SUBAPPLICATION Input_CLIENT_Method_IE (* logiBUS-Taster (logiBUS_IE) loest per CLIENT_0 einen argumentlosen OPC-UA-Methodenaufruf (CALL_METHOD) aus *)
  (* Standard: 61499-2; Description: Copyright (c) 2026 Meisterschulen am Ostbahnhof This program and the accompanying materials are made available under the terms of the Eclipse Public License 2.0 which is available at https://www.eclipse.org/legal/epl-2.0/ SPDX-License-Identifier: EPL-2.0 *)
  (* Version 1.1, 2026-10-18, Franz Höpfinger, Meisterschulen am Ostbahnhof, Wie Button_CLIENT_Method_IE, aber logiBUS_IE statt Button_IE (Taster statt VT-Button) *)
  (* Version 1.0, 2026-09-22, Franz Höpfinger, Meisterschulen am Ostbahnhof, initial implementation - herausgeloest aus logiBUS_AI_Calibrated_Subscribe_VT_OPC (Button_IE + CLIENT_0 kam dort 2x identisch vor, fuer CO und CS). Franz: 'Button_IE CLIENT_0 kann eine Subapp werden, das ist ein generelles Muster zum Rufen einer Methode vom VT aus' - InputEvent ist Parameter (nicht hartcodiert auf BT_PRESSED_LATCHED), damit auch andere Aktivierungsarten (z.B. Loslassen) wiederverwendbar sind. *)
  PACKAGE MyLib::sys;
  IMPORT logiBUS::io::DI::logiBUS_DI;
  IMPORT logiBUS::io::DI::logiBUS_DI_S;
  IMPORT logiBUS::io::DI::logiBUS_DI_Events_S;
  IMPORT logiBUS::io::DI::logiBUS_DI_Events::BUTTON_PRESS_DOWN;
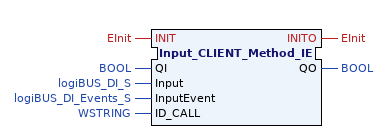
  EVENT_INPUT
    INIT : EInit; (* Initialization Request *)
  END_EVENT
  EVENT_OUTPUT
    INITO : EInit; (* Initialization Confirm *)
  END_EVENT
  VAR_INPUT
    QI : BOOL := TRUE; (* Quality Input - TRUE to enable service *)
    Input : logiBUS::io::DI::logiBUS_DI_S := logiBUS_DI::Invalid; (* Taster Input_I1..I8 *)
    InputEvent : logiBUS::io::DI::logiBUS_DI_Events_S := BUTTON_PRESS_DOWN; (* Welches Tasterereignis den Aufruf ausloest *)
    ID_CALL : WSTRING; (* Methodenadresse (ACTION=CALL_METHOD, mit Endpunkt, auch localhost) *)
  END_VAR
  VAR_OUTPUT
    QO : BOOL; (* Quality Output - TRUE if service executed successfully *)
  END_VAR
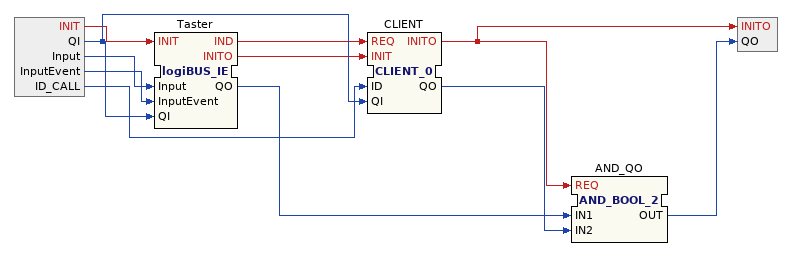
  FBS
    Taster : logiBUS::io::DI::logiBUS_IE;
    CLIENT : iec61499::net::CLIENT_0;
    AND_QO : iec61131::booleanOperators::AND_BOOL_2;
  END_FBS
  EVENT_CONNECTIONS
    Taster.IND TO CLIENT.REQ;
    INIT TO Taster.INIT;
    Taster.INITO TO CLIENT.INIT;
    CLIENT.INITO TO INITO;
    CLIENT.INITO TO AND_QO.REQ;
  END_CONNECTIONS
  DATA_CONNECTIONS
    Input TO Taster.Input;
    InputEvent TO Taster.InputEvent;
    ID_CALL TO CLIENT.ID;
    QI TO Taster.QI;
    QI TO CLIENT.QI;
    Taster.QO TO AND_QO.IN1;
    CLIENT.QO TO AND_QO.IN2;
    AND_QO.OUT TO QO;
  END_CONNECTIONS
END_SUBAPPLICATION
